// TIA Portal project "CMoLibrary_Dev" (V20)

(* hardware
DEVICE "S7-1500/ET200MP station_1"  S7-1500 station
   slot 0: "Rail_0"  Rack  6ES7 590-1***0-0AA0
   slot 1: "PLC_1"  CPU 1516-3 PN/DP  6ES7 516-3AN00-0AB0  V1.8
      slot 3: "CPU display_1"  6ES7591-1BA00-0AA0
      slot 32768: "PROFINET interface_1"  X1
         slot 32769: "Port_1"  X1 P1
         slot 32770: "Port_2"  X1 P2
      slot 33024: "PROFINET interface_2"  X2
         slot 33025: "Port_1"  X2 P1
      slot 33280: "DP interface_1"  X3
*)

// ===== PLC "PLC_1"  CPU 1516-3 PN/DP =====

TYPE "CMoDateTime"
   STRUCT
      RawDateTime : Array[0..6] of DInt;   // Platform-native wall clock data
      Year : DInt := 0;
      Month : DInt := 0;   // 1-12
      Day : DInt := 0;   // 1-31
      Hour : DInt := 0;   // 0-23
      Minute : DInt := 0;   // 0-59
      Second : DInt := 0;   // 0-59
      MicroSecond : DInt := 0;   // 0-999999
      IsLocal : Bool := false;   // TRUE = local time, FALSE = UTC
   END_STRUCT;
END_TYPE

TYPE "CMoDateTimeString"
   STRUCT
      TimeString : String[16];   // HH:MM:SS
      DateString : String[16];   // YYYY-MM-DD
      HMIString : String[32];   // YYYY-MM-DD HH:MM:SS
   END_STRUCT;
END_TYPE

TYPE "CMoHALDigitalInput"
   STRUCT
      Input : Bool := false;   // Raw hardware input (written by device driver)
      QualityInput : Bool := false;   // Hardware health from module status (TRUE = good)
      SimInput : Bool := false;   // Simulation input (written by twin/test)
      EnableSimulation : Bool := false;   // Enable simulation for this point
      SimulationIsActive : Bool := false;   // Computed: EnableSimulation AND Framework.SimulationEnabled
      HandValue : Bool := false;   // Manual override value (set from HMI)
      EnableHand : Bool := false;   // Enable hand mode for this point
      HandIsActive : Bool := false;   // Computed: EnableHand AND Framework.MaintenanceEnabled
      Value : Bool := false;   // THE OUTPUT: conditioned, filtered, mode-selected result
      Inverted : Bool := false;   // Invert input polarity
      BadQualityValue : Bool := false;   // Value to use when quality is bad (safe state)
      EnableDelay : Bool := false;   // Enable debounce filtering
      IsSpare : Bool := false;   // Mark as spare (bypasses quality, forces sim)
      InFilterOnTimeMsec : DInt := 0;   // On-delay debounce (milliseconds)
      InFilterOffTimeMsec : DInt := 0;   // Off-delay debounce (milliseconds)
      PointQuality : Bool := false;   // Computed quality (good if hw OK or sim active)
      RisingEdge : Bool := false;   // One-shot pulse on Value 0 to 1
      FallingEdge : Bool := false;   // One-shot pulse on Value 1 to 0
      "Name" : String[28];   // Human-readable tag name for HMI display
   END_STRUCT;
END_TYPE

TYPE "CMoHALDigitalOutput"
   STRUCT
      Output : Bool := false;   // Physical output (written by FB to hardware)
      QualityInput : Bool := false;   // Hardware health (TRUE = good)
      SimOutput : Bool := false;   // Shadow output for twin consumption during sim
      EnableSimulation : Bool := false;   // Enable simulation for this point
      SimulationIsActive : Bool := false;   // Computed: EnableSimulation AND Framework.SimulationEnabled
      HandValue : Bool := false;   // Manual override value (set from HMI)
      EnableHand : Bool := false;   // Enable hand mode for this point
      HandIsActive : Bool := false;   // Computed: EnableHand AND Framework.MaintenanceEnabled
      Value : Bool := false;   // Business logic command
      Inverted : Bool := false;   // Invert output polarity
      BadQualityValue : Bool := false;   // Value when quality is bad (safe state)
      IsSpare : Bool := false;   // Mark as spare
      PointQuality : Bool := false;   // Computed quality
      "Name" : String[28];   // Human-readable tag name
   END_STRUCT;
END_TYPE

TYPE "CMoInterlock"
   STRUCT
      PointCount : Int := 4;   // Number of active conditions (1-16)
      Condition : Array[0..15] of Bool;   // Condition inputs (set by business logic each scan)
      Bypass : Array[0..15] of Bool;   // Per-condition bypass (set from HMI)
      OK : Bool := false;   // All active conditions met (or bypassed)
      InBypass : Bool := false;   // At least one condition is bypassed
      BypassAlarm : Bool := false;   // Alarm: operating with bypassed conditions
      FirstOut : Int := -1;   // Index of first condition to drop (-1 = none)
      ConditionMet : Array[0..15] of Bool;   // Condition OR its bypass
      ConditionFaulted : Array[0..15] of Bool;   // Failed AND not bypassed
      "Name" : String[28];   // Interlock name
      ConditionName : Array[0..15] of String[28];   // Per-condition labels
   END_STRUCT;
END_TYPE

TYPE "CMoFramework"
   STRUCT
      AnyAudibleOn : Bool := false;   // At least one alarm has audible active
      AnyAudibleOnLastScan : Bool := false;   // Scratch accumulator
      AnyAlarmActive : Bool := false;   // At least one alarm active
      AnyAlarmActiveLastScan : Bool := false;   // Scratch accumulator
      AnyWarningActive : Bool := false;   // At least one warning-severity alarm
      AnyWarningActiveLastScan : Bool := false;   // Scratch accumulator
      AnyFaultActive : Bool := false;   // At least one fault-severity alarm
      AnyFaultActiveLastScan : Bool := false;   // Scratch accumulator
      AnyCriticalActive : Bool := false;   // At least one critical-severity alarm
      AnyCriticalActiveLastScan : Bool := false;   // Scratch accumulator
      AnySimulationOn : Bool := false;   // At least one I/O in simulation mode
      AnySimulationOnLastScan : Bool := false;   // Scratch accumulator
      AnyHandOn : Bool := false;   // At least one I/O in hand mode
      AnyHandOnLastScan : Bool := false;   // Scratch accumulator
      SilenceCmd : Bool := false;   // HMI silence button (momentary)
      GlobalAlmRstCmd : Bool := false;   // HMI global alarm reset (momentary)
      GlobalAlmRstEn : Bool := false;   // Enable global alarm reset
      SimulationEnabled : Bool := false;   // Master simulation enable
      EmulationEnabled : Bool := false;   // Running on emulated controller
      MaintenanceEnabled : Bool := false;   // Enables Hand mode
      Tick100ms : Bool := false;   // Pulse TRUE for one scan every 100ms
      Tick1s : Bool := false;   // Pulse TRUE for one scan every 1s
      Tick10s : Bool := false;   // Pulse TRUE for one scan every 10s
      Blink100ms : Bool := false;   // 100ms on/off blinker
      Blink250ms : Bool := false;   // 250ms on/off blinker
      Blink500ms : Bool := false;   // 500ms on/off blinker
      Blink1s : Bool := false;   // 1s on/off blinker
      Blink2s : Bool := false;   // 2s on/off blinker
      InhibitAlarms : Bool := false;   // Corporate alarm inhibit
      AlwaysTrue : Bool := false;   // Constant TRUE
      AlwaysFalse : Bool := false;   // Constant FALSE
      ApplicationCount : DInt := 0;   // Number of AOI instances registered
      AlarmCount : Int := 0;   // Current active alarm count
      TempAlarmCount : Int := 0;   // Scratch accumulator
      FreeRunningTimer : DInt := 0;   // Free-running ms counter
      LastRandomSeed : DInt := 0;   // Seed for random number generator
      Random : Real := 0.0;   // Current random number 0.0-1.0
      CycleTime : Real := 0.0;   // Last scan time (milliseconds)
      InhibitAlarmGroups : Array[0..15] of DWord;   // Per-group alarm inhibit (512 groups)
      CurrentUTCDateTime : "CMoDateTime";   // Current UTC time
      CurrentLocalDateTime : "CMoDateTime";   // Current local time
      CurrentUTCString : "CMoDateTimeString";   // UTC time formatted strings
      CurrentLocalString : "CMoDateTimeString";   // Local time formatted strings
      NotUsedDI : "CMoHALDigitalInput";   // Spare DI HAL instance
      NotUsedDO : "CMoHALDigitalOutput";   // Spare DO HAL instance
      ModuleStatusMinInterval : DInt := 5000;   // ms between module checks
      ModuleStatusRandomDistribution : DInt := 2000;   // ms random spread for check timing
      ModuleStatusGraceTime : DInt := 30000;   // ms before declaring module lost
   END_STRUCT;
END_TYPE

DATA_BLOCK "GVL"   // DB1
{ S7_Optimized_Access := 'TRUE' }
VERSION : 0.1
   VAR
      Framework : "CMoFramework";
      DI_PartPresent : "CMoHALDigitalInput";
      DI_GuardClosed : "CMoHALDigitalInput";
      DO_MotorRun : "CMoHALDigitalOutput";
      Interlock_Motor : "CMoInterlock";
      SimPartPresent : Bool;
      SimGuardClosed : Bool;
      saveStart : Bool;
      startDate : "CMoDateTime";
      saveEnd : Bool;
      endDate : "CMoDateTime";
   END_VAR
BEGIN
END_DATA_BLOCK

DATA_BLOCK "fbGuardClosed"   // DB2
{ S7_Optimized_Access := 'TRUE' }
VERSION : 0.1
// stored: InstanceOfName CMoDigitalInput
"CMoDigitalInput"
BEGIN
END_DATA_BLOCK

DATA_BLOCK "fbInterlock"   // DB3
{ S7_Optimized_Access := 'TRUE' }
VERSION : 0.1
// stored: InstanceOfName CMoEvalInterlock
"CMoEvalInterlock"
BEGIN
END_DATA_BLOCK

DATA_BLOCK "fbPartPresent"   // DB4
{ S7_Optimized_Access := 'TRUE' }
VERSION : 0.1
// stored: InstanceOfName CMoDigitalInput
"CMoDigitalInput"
BEGIN
END_DATA_BLOCK

DATA_BLOCK "fbMainRoutine"   // DB5
{ S7_Optimized_Access := 'TRUE' }
VERSION : 0.1
// stored: InstanceOfName CMoMainRuntime
"CMoMainRuntime"
BEGIN
END_DATA_BLOCK

DATA_BLOCK "fbMotorRun"   // DB6
{ S7_Optimized_Access := 'TRUE' }
VERSION : 0.1
// stored: InstanceOfName CMoDigitalOutput
"CMoDigitalOutput"
BEGIN
END_DATA_BLOCK

DATA_BLOCK "CMoDiffTime_DB"   // DB7
{ S7_Optimized_Access := 'TRUE' }
VERSION : 0.1
// stored: InstanceOfName CMoDiffTime
"CMoDiffTime"
BEGIN
END_DATA_BLOCK

FUNCTION_BLOCK "CMoRandom"   // FB1, SCL
{ S7_Optimized_Access := 'TRUE' }
VERSION : 0.1
   VAR_INPUT
      Seed : DInt := 48271;
   END_VAR
   VAR_OUTPUT
      Out : Real;
      NewSeed : DInt;
   END_VAR
BEGIN

   // =============================================================================
   // CMoRandom â€” Random Number Generator
   // CMo Library v1.0
   // =============================================================================
   // Park-Miller linear congruential generator.
   // Outputs a REAL between 0.0 and 1.0.
   //
   // Feed Seed from Framework.LastRandomSeed, write NewSeed back after call.
   // Called internally by CMoMainRuntime every scan.
   //
   // Usage:
   //   fbRandom(Seed := Framework.LastRandomSeed);
   //   Framework.Random := fbRandom.Out;
   //   Framework.LastRandomSeed := fbRandom.NewSeed;
   // =============================================================================

   // Ensure positive seed
   IF #Seed <= 0 THEN
       #Seed := 1;
   END_IF;

   // Park-Miller LCG: next = (seed * 16807) MOD 2147483647
   #NewSeed := (#Seed MOD 127773) * 16807 - (#Seed / 127773) * 2836;
   IF #NewSeed <= 0 THEN
       #NewSeed := #NewSeed + 2147483647;
   END_IF;

   #Out := DINT_TO_REAL(#NewSeed) / 2147483647.0;
END_FUNCTION_BLOCK

FUNCTION_BLOCK "CMoGetLocalDateTime"   // FB2, SCL
{ S7_Optimized_Access := 'TRUE' }
VERSION : 0.1
   VAR_IN_OUT
      DateTime : "CMoDateTime";
   END_VAR
   VAR_TEMP
      dtlNow : DTL;
      retVal : Int;
   END_VAR
BEGIN

   // =============================================================================
   // CMoGetLocalDateTime â€” Read Local System Time (Siemens)
   // CMo Library v1.0
   // =============================================================================
   // Reads the local system time using RD_LOC_T and parses DTL fields
   // into CMoDateTime.
   //
   // Must be called cyclically. Called internally by CMoMainRuntime.
   //
   // Usage:
   //   fbLocal(DateTime := Framework.CurrentLocalDateTime);
   // =============================================================================

   #retVal := RD_LOC_T(#dtlNow);

   IF #retVal <= 1 THEN
       #DateTime.Year := INT_TO_DINT(#dtlNow.YEAR);
       #DateTime.Month := USINT_TO_DINT(#dtlNow.MONTH);
       #DateTime.Day := USINT_TO_DINT(#dtlNow.DAY);
       #DateTime.Hour := USINT_TO_DINT(#dtlNow.HOUR);
       #DateTime.Minute := USINT_TO_DINT(#dtlNow.MINUTE);
       #DateTime.Second := USINT_TO_DINT(#dtlNow.SECOND);
       #DateTime.MicroSecond := UDINT_TO_DINT(#dtlNow.NANOSECOND / 1000);
       #DateTime.IsLocal := TRUE;
   END_IF;
END_FUNCTION_BLOCK

FUNCTION_BLOCK "CMoGetUTCDateTime"   // FB3, SCL
{ S7_Optimized_Access := 'TRUE' }
VERSION : 0.1
   VAR_IN_OUT
      DateTime : "CMoDateTime";
   END_VAR
   VAR_TEMP
      dtlNow : DTL;
      retVal : Int;
   END_VAR
BEGIN

   // =============================================================================
   // CMoGetUTCDateTime â€” Read UTC System Time (Siemens)
   // CMo Library v1.0
   // =============================================================================
   // Reads the UTC system time using RD_SYS_T and parses DTL fields
   // into CMoDateTime.
   //
   // RD_SYS_T returns UTC on S7-1500.
   // Must be called cyclically. Called internally by CMoMainRuntime.
   //
   // Usage:
   //   fbUTC(DateTime := Framework.CurrentUTCDateTime);
   // =============================================================================

   #retVal := RD_SYS_T(#dtlNow);

   IF #retVal = 0 THEN
       #DateTime.Year := INT_TO_DINT(#dtlNow.YEAR);
       #DateTime.Month := USINT_TO_DINT(#dtlNow.MONTH);
       #DateTime.Day := USINT_TO_DINT(#dtlNow.DAY);
       #DateTime.Hour := USINT_TO_DINT(#dtlNow.HOUR);
       #DateTime.Minute := USINT_TO_DINT(#dtlNow.MINUTE);
       #DateTime.Second := USINT_TO_DINT(#dtlNow.SECOND);
       #DateTime.MicroSecond := UDINT_TO_DINT(#dtlNow.NANOSECOND / 1000);
       #DateTime.IsLocal := FALSE;
   END_IF;
END_FUNCTION_BLOCK

FUNCTION_BLOCK "CMoElapsedTime"   // FB4, SCL
{ S7_Optimized_Access := 'TRUE' }
VERSION : 0.1
   VAR_INPUT
      Start : Bool;
      Stop : Bool;
      Reset : Bool;
   END_VAR
   VAR_OUTPUT
      ElapsedMs : Real;
      Running : Bool;
   END_VAR
   VAR
      PrevStart : Bool;
      PrevStop : Bool;
      tmRun : TON_TIME;
      Capturing : Bool;
   END_VAR
BEGIN

   // =============================================================================
   // CMoElapsedTime â€” Elapsed Time Measurement
   // CMo Library v1.0
   // =============================================================================
   // Measures elapsed time between Start and Stop rising edges.
   // Uses a TON timer internally for millisecond-resolution measurement.
   // Live readout available via ElapsedMs while Running is TRUE.
   //
   // Usage:
   //   myTimer(Start := TRUE);       // Begin measurement
   //   // ... code or scans pass ...
   //   myTimer(Stop := TRUE);        // End measurement
   //   result := myTimer.ElapsedMs;  // Read duration in ms
   //   myTimer(Reset := TRUE);       // Clear for next use
   // =============================================================================

   // Reset: clear everything
   IF #Reset THEN
       #ElapsedMs := 0.0;
       #Running := FALSE;
       #Capturing := FALSE;
       RETURN;
   END_IF;

   // Start on rising edge
   IF #Start AND NOT #PrevStart THEN
       #Capturing := TRUE;
       #Running := TRUE;
       #tmRun(IN := FALSE,
              PT := T#24D);
   END_IF;
   #PrevStart := #Start;

   // Accumulate while running
   IF #Capturing THEN
       #tmRun(IN := TRUE,
              PT := T#24D);
       #ElapsedMs := DINT_TO_REAL(TIME_TO_DINT(#tmRun.ET));
   END_IF;

   // Stop on rising edge
   IF #Stop AND NOT #PrevStop AND #Capturing THEN
       #ElapsedMs := DINT_TO_REAL(TIME_TO_DINT(#tmRun.ET));
       #Capturing := FALSE;
       #Running := FALSE;
   END_IF;
   #PrevStop := #Stop;
END_FUNCTION_BLOCK

FUNCTION_BLOCK "CMoDateTimeToString"   // FB5, SCL
{ S7_Optimized_Access := 'TRUE' }
VERSION : 0.1
   VAR_INPUT
      DateTime : "CMoDateTime";
   END_VAR
   VAR_IN_OUT
      DateTimeString : "CMoDateTimeString";
   END_VAR
   VAR_TEMP
      sYear : String[5];
      sMonth : String[3];
      sDay : String[3];
      sHour : String[3];
      sMinute : String[3];
      sSecond : String[3];
      sTemp : String[40];
   END_VAR
BEGIN
   // =============================================================================
   // CMoDateTimeToString — Format DateTime for HMI Display
   // CMo Library v1.0
   // =============================================================================
   // Converts CMoDateTime fields into zero-padded human-readable strings:
   //   TimeString: "HH:MM:SS"
   //   DateString: "YYYY-MM-DD"
   //   HMIString:  "YYYY-MM-DD HH:MM:SS"
   //
   // Siemens DINT_TO_STRING prepends a '+' sign. DELETE strips it.
   //
   // Usage:
   //   fbFmt(DateTime := myTime, DateTimeString := myStrings);
   // =============================================================================

   // Convert and strip leading '+'
   #sYear := DELETE(IN := DINT_TO_STRING(#DateTime.Year), L := 1, P := 1);

   IF #DateTime.Month < 10 THEN
       #sMonth := CONCAT(IN1 := '0', IN2 := DELETE(IN := DINT_TO_STRING(#DateTime.Month), L := 1, P := 1));
   ELSE
       #sMonth := DELETE(IN := DINT_TO_STRING(#DateTime.Month), L := 1, P := 1);
   END_IF;

   IF #DateTime.Day < 10 THEN
       #sDay := CONCAT(IN1 := '0', IN2 := DELETE(IN := DINT_TO_STRING(#DateTime.Day), L := 1, P := 1));
   ELSE
       #sDay := DELETE(IN := DINT_TO_STRING(#DateTime.Day), L := 1, P := 1);
   END_IF;

   IF #DateTime.Hour < 10 THEN
       #sHour := CONCAT(IN1 := '0', IN2 := DELETE(IN := DINT_TO_STRING(#DateTime.Hour), L := 1, P := 1));
   ELSE
       #sHour := DELETE(IN := DINT_TO_STRING(#DateTime.Hour), L := 1, P := 1);
   END_IF;

   IF #DateTime.Minute < 10 THEN
       #sMinute := CONCAT(IN1 := '0', IN2 := DELETE(IN := DINT_TO_STRING(#DateTime.Minute), L := 1, P := 1));
   ELSE
       #sMinute := DELETE(IN := DINT_TO_STRING(#DateTime.Minute), L := 1, P := 1);
   END_IF;

   IF #DateTime.Second < 10 THEN
       #sSecond := CONCAT(IN1 := '0', IN2 := DELETE(IN := DINT_TO_STRING(#DateTime.Second), L := 1, P := 1));
   ELSE
       #sSecond := DELETE(IN := DINT_TO_STRING(#DateTime.Second), L := 1, P := 1);
   END_IF;

   // Build TimeString: "HH:MM:SS"
   #sTemp := CONCAT(IN1 := #sHour, IN2 := ':');
   #sTemp := CONCAT(IN1 := #sTemp, IN2 := #sMinute);
   #sTemp := CONCAT(IN1 := #sTemp, IN2 := ':');
   #sTemp := CONCAT(IN1 := #sTemp, IN2 := #sSecond);
   #DateTimeString.TimeString := #sTemp;

   // Build DateString: "YYYY-MM-DD"
   #sTemp := CONCAT(IN1 := #sYear, IN2 := '-');
   #sTemp := CONCAT(IN1 := #sTemp, IN2 := #sMonth);
   #sTemp := CONCAT(IN1 := #sTemp, IN2 := '-');
   #sTemp := CONCAT(IN1 := #sTemp, IN2 := #sDay);
   #DateTimeString.DateString := #sTemp;

   // Build HMIString: "YYYY-MM-DD HH:MM:SS"
   #sTemp := CONCAT(IN1 := #DateTimeString.DateString, IN2 := ' ');
   #sTemp := CONCAT(IN1 := #sTemp, IN2 := #DateTimeString.TimeString);
   #DateTimeString.HMIString := #sTemp;
END_FUNCTION_BLOCK

FUNCTION_BLOCK "CMoDiffTime"   // FB6, SCL
{ S7_Optimized_Access := 'TRUE' }
VERSION : 0.1
   VAR_INPUT
      StartTime : "CMoDateTime";
      EndTime : "CMoDateTime";
   END_VAR
   VAR_OUTPUT
      Result : "CMoDateTime";
      TotalSeconds : DInt;
      TotalMicroseconds : DInt;
   END_VAR
   VAR_TEMP
      Borrow : DInt;
      Diff : DInt;
      "a" : DInt;
      y : DInt;
      "m" : DInt;
      jdnStart : DInt;
      jdnEnd : DInt;
      diffDays : DInt;
      diffUs : DInt;
      diffSec : DInt;
      diffMin : DInt;
      diffHr : DInt;
   END_VAR
BEGIN
   // =============================================================================
   // CMoDiffTime — DateTime Subtraction via Julian Day Number
   // CMo Library v1.0
   // =============================================================================
   // Computes (EndTime - StartTime) using Julian Day Number conversion.
   // Converts both dates to JDN (integer day count), subtracts, then
   // handles sub-day time remainder with borrow propagation.
   //
   // This is mathematically correct for all valid dates regardless of
   // month lengths, leap years, or century boundaries.
   //
   // Usage:
   //   fbDiff(StartTime := tStart, EndTime := tEnd);
   //   elapsed := fbDiff.TotalSeconds;
   // =============================================================================

   // JDN for StartTime
   #a := (14 - #StartTime.Month) / 12;
   #y := #StartTime.Year + 4800 - #a;
   #m := #StartTime.Month + 12 * #a - 3;
   #jdnStart := #StartTime.Day + (153 * #m + 2) / 5 + 365 * #y + #y / 4 - #y / 100 + #y / 400 - 32045;

   // JDN for EndTime
   #a := (14 - #EndTime.Month) / 12;
   #y := #EndTime.Year + 4800 - #a;
   #m := #EndTime.Month + 12 * #a - 3;
   #jdnEnd := #EndTime.Day + (153 * #m + 2) / 5 + 365 * #y + #y / 4 - #y / 100 + #y / 400 - 32045;

   // Day difference
   #diffDays := #jdnEnd - #jdnStart;

   // Sub-day difference with borrow propagation
   #diffUs := #EndTime.MicroSecond - #StartTime.MicroSecond;
   IF #diffUs < 0 THEN
       #diffUs := #diffUs + 1000000;
       #diffSec := -1;
   ELSE
       #diffSec := 0;
   END_IF;

   #diffSec := #diffSec + #EndTime.Second - #StartTime.Second;
   IF #diffSec < 0 THEN
       #diffSec := #diffSec + 60;
       #diffMin := -1;
   ELSE
       #diffMin := 0;
   END_IF;

   #diffMin := #diffMin + #EndTime.Minute - #StartTime.Minute;
   IF #diffMin < 0 THEN
       #diffMin := #diffMin + 60;
       #diffHr := -1;
   ELSE
       #diffHr := 0;
   END_IF;

   #diffHr := #diffHr + #EndTime.Hour - #StartTime.Hour;
   IF #diffHr < 0 THEN
       #diffHr := #diffHr + 24;
       #diffDays := #diffDays - 1;
   END_IF;

   // Populate result
   #Result.Year := 0;
   #Result.Month := 0;
   #Result.Day := #diffDays;
   #Result.Hour := #diffHr;
   #Result.Minute := #diffMin;
   #Result.Second := #diffSec;
   #Result.MicroSecond := #diffUs;
   #Result.IsLocal := FALSE;

   // Convenience totals
   #TotalSeconds := #diffSec + (#diffMin * 60) + (#diffHr * 3600) + (#diffDays * 86400);
   #TotalMicroseconds := #diffUs;
END_FUNCTION_BLOCK

FUNCTION_BLOCK "CMoAlarm"   // FB7, SCL
{ S7_Optimized_Access := 'TRUE' }
VERSION : 0.1
   VAR_INPUT
      Trigger : Bool;
      EnableAlarm : Bool := TRUE;
      AlarmOnTrue : Bool := TRUE;
      AutoReset : Bool;
      Delay : DInt;
      GroupNo : DInt;
      ID : Int;
      IsWarning : Bool;
      IsFault : Bool;
      IsCritical : Bool;
      EnableAudio : Bool;
      SystemResetEnable : Bool := TRUE;
      Inhibit : Bool;
      CountPreset : DInt;
   END_VAR
   VAR_OUTPUT
      AlarmActive : Bool;
      InhibitActive : Bool;
      AlarmCount : DInt;
      CountExceeded : Bool;
      AlarmSilenced : Bool;
   END_VAR
   VAR_IN_OUT
      Framework : "CMoFramework";
      CountReset : Bool;
      Reset : Bool;
   END_VAR
   VAR
      AlarmTimer : TON_TIME;
      IntGroupNo : DInt;
      IntID : DInt;
      IntReset : Bool;
      TriggerCondition : Bool;
      PrevAlarmActive : Bool;
      GroupWord : DInt;
      GroupBit : DInt;
   END_VAR
BEGIN

   // =============================================================================
   // CMoAlarm â€” Alarm Monitor
   // CMo Library v1.0
   // =============================================================================
   // Monitors a trigger condition and manages alarm lifecycle.
   // Supports configurable trigger polarity, delay before activation,
   // auto/manual reset, occurrence counting with threshold,
   // severity classification (Warning/Fault/Critical), group-based
   // inhibit, and HMI silencing.
   //
   // Usage:
   //   fbAlarm(
   //       Framework := GVL.Framework,
   //       Trigger := SomeCondition,
   //       ID := 100,
   //       Delay := 2000,
   //       IsFault := TRUE
   //   );
   // =============================================================================

   // Clamp group and ID
   IF #GroupNo >= 0 AND #GroupNo <= 511 THEN
       #IntGroupNo := #GroupNo;
   ELSE
       #IntGroupNo := 0;
   END_IF;

   IF #ID >= 1 AND #ID <= 9023 THEN
       #IntID := #ID;
   ELSE
       #IntID := 0;
   END_IF;

   #GroupWord := #IntGroupNo / 32;
   #GroupBit := #IntGroupNo MOD 32;

   // Count reset
   IF #CountReset THEN
       #AlarmCount := 0;
       #CountReset := FALSE;
   END_IF;

   // Inhibit evaluation
   #InhibitActive := NOT #EnableAlarm
   OR #Inhibit
   OR #Framework.InhibitAlarms;
   IF NOT #InhibitActive AND (#Framework.InhibitAlarmGroups[#GroupWord] AND SHL(IN := DWORD#1, N := DINT_TO_INT(#GroupBit))) <> 0 THEN
       #InhibitActive := TRUE;
   END_IF;

   // Composite reset
   #IntReset := #AutoReset
   OR #Reset
   OR (#SystemResetEnable AND #Framework.GlobalAlmRstEn AND #Framework.GlobalAlmRstCmd);

   // Trigger polarity
   IF #AlarmOnTrue THEN
       #TriggerCondition := #Trigger;
   ELSE
       #TriggerCondition := NOT #Trigger;
   END_IF;

   // Alarm activation with delay
   IF #IntID <> 0 THEN
       #AlarmTimer(
                   IN := (NOT #InhibitActive AND #TriggerCondition) OR (#AlarmActive AND NOT #IntReset),
                   PT := DINT_TO_TIME(#Delay)
       );
       #AlarmActive := #AlarmTimer.Q;
   ELSE
       #AlarmActive := FALSE;
   END_IF;

   // Count activations (rising edge)
   IF #AlarmActive AND NOT #PrevAlarmActive THEN
       #AlarmCount := #AlarmCount + 1;
   END_IF;

   // Silence
   IF #AlarmActive THEN
       IF #Framework.SilenceCmd OR #AlarmSilenced THEN
           #AlarmSilenced := TRUE;
       END_IF;
   ELSE
       #AlarmSilenced := FALSE;
   END_IF;

   // Roll up into Framework
   IF #AlarmActive THEN
       #Framework.TempAlarmCount := #Framework.TempAlarmCount + 1;
       #Framework.AnyAlarmActiveLastScan := TRUE;

       IF NOT #AlarmSilenced THEN
           IF #EnableAudio THEN
               #Framework.AnyAudibleOnLastScan := TRUE;
           END_IF;
           IF #IsWarning THEN
               #Framework.AnyWarningActiveLastScan := TRUE;
           END_IF;
           IF #IsFault THEN
               #Framework.AnyFaultActiveLastScan := TRUE;
           END_IF;
           IF #IsCritical THEN
               #Framework.AnyCriticalActiveLastScan := TRUE;
           END_IF;
       END_IF;
   END_IF;

   // Count threshold
   #CountExceeded := (#CountPreset > 0) AND (#AlarmCount >= #CountPreset);

   // Clear manual reset
   #Reset := FALSE;

   // Previous state
   #PrevAlarmActive := #AlarmActive;
END_FUNCTION_BLOCK

FUNCTION_BLOCK "CMoDigitalInput"   // FB8, SCL
{ S7_Optimized_Access := 'TRUE' }
VERSION : 0.1
   VAR_INPUT
      DeviceInput : Bool;
      QualityInput : Bool;
   END_VAR
   VAR_IN_OUT
      HAL : "CMoHALDigitalInput";
      Framework : "CMoFramework";
   END_VAR
   VAR
      ConditionedInput : Bool;
      DebouncedValue : Bool;
      OnDelayTimer : TON_TIME;
      OffDelayTimer : TOF_TIME;
      PrevValue : Bool;
      FirstScan : Bool := TRUE;
      ReSync : Bool;
      NoFilterNeeded : Bool;
   END_VAR
BEGIN

   // =============================================================================
   // CMoDigitalInput â€” Digital Input Signal Conditioning
   // CMo Library v1.0
   // =============================================================================
   // Takes a raw hardware input and produces a conditioned .Value through:
   //   1. Mode determination (Normal / Simulation / Hand)
   //   2. Quality evaluation (hardware health, sim, spare)
   //   3. Mode selection + polarity inversion
   //   4. Debounce filtering (configurable on/off delay with resync)
   //   5. Hand value bumpless transfer
   //   6. Quality gating (bad quality -> configurable fallback)
   //   7. Edge detection (RisingEdge / FallingEdge one-shot pulses)
   //
   // Business logic reads .Value only. Never touch .Input, .SimInput,
   // .HandValue, or any plumbing directly.
   //
   // Usage:
   //   fbInput(
   //       HAL := GVL.MyInput,
   //       DeviceInput := Module1:I.Data[0],
   //       QualityInput := Module1_Status.Running,
   //       Framework := GVL.Framework
   //   );
   // =============================================================================

   // Mode determination
   #HAL.HandIsActive := #HAL.EnableHand AND #Framework.MaintenanceEnabled;
   IF #HAL.HandIsActive THEN
       #Framework.AnyHandOnLastScan := TRUE;
   END_IF;

   #HAL.SimulationIsActive := #HAL.EnableSimulation AND #Framework.SimulationEnabled;
   IF #HAL.SimulationIsActive THEN
       #Framework.AnySimulationOnLastScan := TRUE;
   END_IF;

   // Point quality
   IF #HAL.IsSpare THEN
       #HAL.PointQuality := TRUE;
   ELSIF #HAL.SimulationIsActive THEN
       #HAL.PointQuality := TRUE;
   ELSE
       #HAL.QualityInput := #QualityInput;
       #HAL.PointQuality := #QualityInput;
   END_IF;

   // Latch raw input
   #HAL.Input := #DeviceInput;

   // Mode selection + inversion
   IF #HAL.SimulationIsActive THEN
       IF #HAL.Inverted THEN
           #ConditionedInput := NOT #HAL.SimInput;
       ELSE
           #ConditionedInput := #HAL.SimInput;
       END_IF;
   ELSE
       IF #HAL.Inverted THEN
           #ConditionedInput := NOT #HAL.Input;
       ELSE
           #ConditionedInput := #HAL.Input;
       END_IF;
   END_IF;

   // Debounce filter
   IF NOT #HAL.EnableDelay THEN
       #DebouncedValue := #ConditionedInput;
       #ReSync := TRUE;
   ELSE
       IF #HAL.InFilterOnTimeMsec < 0 THEN
           #HAL.InFilterOnTimeMsec := 0;
       END_IF;
       IF #HAL.InFilterOffTimeMsec < 0 THEN
           #HAL.InFilterOffTimeMsec := 0;
       END_IF;

       #OnDelayTimer(
                     IN := #ConditionedInput OR (#OffDelayTimer.Q AND #OnDelayTimer.Q),
                     PT := DINT_TO_TIME(#HAL.InFilterOnTimeMsec)
       );

       #OffDelayTimer(
                      IN := #ConditionedInput,
                      PT := DINT_TO_TIME(#HAL.InFilterOffTimeMsec)
       );

       #NoFilterNeeded := (#ConditionedInput AND #OnDelayTimer.Q)
       OR (NOT #ConditionedInput AND NOT #OffDelayTimer.Q);

       IF #ReSync THEN
           IF (#DebouncedValue AND #OnDelayTimer.Q) OR
               (NOT #DebouncedValue AND NOT #OnDelayTimer.Q) THEN
               #ReSync := FALSE;
           END_IF;
       END_IF;

       IF #ReSync OR #HAL.IsSpare THEN
           #DebouncedValue := #ConditionedInput;
       ELSIF #OnDelayTimer.Q THEN
           #DebouncedValue := TRUE;
       ELSIF NOT #OffDelayTimer.Q THEN
           #DebouncedValue := FALSE;
       END_IF;
   END_IF;

   // Hand value tracking (bumpless transfer)
   IF NOT #HAL.HandIsActive THEN
       #HAL.HandValue := #HAL.Value;
   END_IF;

   // Final value with quality gating
   IF #HAL.PointQuality THEN
       IF #HAL.HandIsActive THEN
           #HAL.Value := #HAL.HandValue;
       ELSE
           #HAL.Value := #DebouncedValue;
       END_IF;
   ELSE
       #HAL.Value := #HAL.BadQualityValue;
   END_IF;

   // Edge detection
   IF #FirstScan THEN
       #PrevValue := #HAL.Value;
       #HAL.RisingEdge := FALSE;
       #HAL.FallingEdge := FALSE;
       #FirstScan := FALSE;
   ELSE
       #HAL.RisingEdge := #HAL.Value AND NOT #PrevValue;
       #HAL.FallingEdge := NOT #HAL.Value AND #PrevValue;
       #PrevValue := #HAL.Value;
   END_IF;
END_FUNCTION_BLOCK

FUNCTION_BLOCK "CMoDigitalOutput"   // FB9, SCL
{ S7_Optimized_Access := 'TRUE' }
VERSION : 0.1
   VAR_INPUT
      QualityInput : Bool;
   END_VAR
   VAR_OUTPUT
      DeviceOutput : Bool;
   END_VAR
   VAR_IN_OUT
      HAL : "CMoHALDigitalOutput";
      Framework : "CMoFramework";
   END_VAR
   VAR
      ConditionedOutput : Bool;
      OutputWithHand : Bool;
   END_VAR
BEGIN

   // =============================================================================
   // CMoDigitalOutput â€” Digital Output Signal Conditioning
   // CMo Library v1.0
   // =============================================================================
   // Takes .Value written by business logic and produces a conditioned
   // physical output through:
   //   1. Mode determination (Normal / Simulation / Hand)
   //   2. Quality evaluation (hardware health, sim, spare)
   //   3. Polarity inversion
   //   4. Hand value bumpless transfer
   //   5. Hand mode selection
   //   6. Simulation gating (suppress physical output, capture to .SimOutput)
   //
   // In simulation mode: DeviceOutput is suppressed. The digital twin
   // reads .SimOutput to see what business logic commanded.
   //
   // Usage:
   //   fbOutput(
   //       HAL := GVL.MyOutput,
   //       QualityInput := Module2_Status.Running,
   //       Framework := GVL.Framework
   //   );
   //   Module2:O.Data[0] := fbOutput.DeviceOutput;
   // =============================================================================

   // Mode determination
   #HAL.HandIsActive := #HAL.EnableHand AND #Framework.MaintenanceEnabled AND NOT #HAL.IsSpare;
   IF #HAL.HandIsActive THEN
       #Framework.AnyHandOnLastScan := TRUE;
   END_IF;

   #HAL.SimulationIsActive := #HAL.EnableSimulation AND #Framework.SimulationEnabled;
   IF #HAL.SimulationIsActive THEN
       #Framework.AnySimulationOnLastScan := TRUE;
   END_IF;

   // Point quality
   IF #HAL.IsSpare THEN
       #HAL.PointQuality := TRUE;
   ELSIF #HAL.SimulationIsActive THEN
       #HAL.PointQuality := TRUE;
   ELSE
       #HAL.QualityInput := #QualityInput;
       #HAL.PointQuality := #QualityInput;
   END_IF;

   // Inversion
   IF NOT #HAL.IsSpare THEN
       IF #HAL.Inverted THEN
           #ConditionedOutput := NOT #HAL.Value;
       ELSE
           #ConditionedOutput := #HAL.Value;
       END_IF;
   ELSE
       #ConditionedOutput := FALSE;
   END_IF;

   // Hand value tracking (bumpless transfer)
   IF NOT #HAL.HandIsActive THEN
       #HAL.HandValue := #HAL.Value;
   END_IF;

   // Hand mode selection
   IF #HAL.HandIsActive THEN
       #OutputWithHand := #HAL.HandValue;
   ELSE
       #OutputWithHand := #ConditionedOutput;
   END_IF;

   // Simulation gating
   IF #HAL.SimulationIsActive THEN
       #DeviceOutput := FALSE;
   ELSE
       #DeviceOutput := #OutputWithHand;
   END_IF;

   #HAL.SimOutput := #OutputWithHand;
   #HAL.Output := #DeviceOutput;
END_FUNCTION_BLOCK

FUNCTION_BLOCK "CMoEvalInterlock"   // FB10, SCL
{ S7_Optimized_Access := 'TRUE' }
VERSION : 0.1
   VAR_IN_OUT
      Ilk : "CMoInterlock";
   END_VAR
   VAR
      PrevOK : Bool;
   END_VAR
   VAR_TEMP
      i : Int;
      AllMet : Bool;
      AnyBypassed : Bool;
      FirstDropped : Int;
   END_VAR
BEGIN

   // =============================================================================
   // CMoEvalInterlock â€” Interlock Evaluation
   // CMo Library v1.0
   // =============================================================================
   // Evaluates up to 16 AND conditions with first-out tracking
   // and per-condition bypass. All active conditions must be TRUE
   // (or bypassed) for .OK to be TRUE.
   //
   // FirstOut latches the index of the first faulted condition on
   // the OK->NOT OK transition (root cause analysis from HMI).
   //
   // Usage:
   //   Ilk.Condition[0] := EStop.Value;
   //   Ilk.Condition[1] := GuardDoor.Value;
   //   fbInterlock(Ilk := MyInterlock);
   //   IF MyInterlock.OK THEN ... END_IF;
   // =============================================================================

   // Clamp PointCount
   IF #Ilk.PointCount < 1 THEN
       #Ilk.PointCount := 1;
   ELSIF #Ilk.PointCount > 16 THEN
       #Ilk.PointCount := 16;
   END_IF;

   // Evaluate each condition
   #AllMet := TRUE;
   #AnyBypassed := FALSE;
   #FirstDropped := -1;

   FOR #i := 0 TO #Ilk.PointCount - 1 DO
       #Ilk.ConditionMet[#i] := #Ilk.Condition[#i] OR #Ilk.Bypass[#i];
       #Ilk.ConditionFaulted[#i] := NOT #Ilk.Condition[#i] AND NOT #Ilk.Bypass[#i];

       IF #Ilk.Bypass[#i] THEN
           #AnyBypassed := TRUE;
       END_IF;

       IF #Ilk.ConditionFaulted[#i] AND #FirstDropped = -1 THEN
           #FirstDropped := #i;
       END_IF;

       IF NOT #Ilk.ConditionMet[#i] THEN
           #AllMet := FALSE;
       END_IF;
   END_FOR;

   // Clear unused conditions
   FOR #i := #Ilk.PointCount TO 15 DO
       #Ilk.ConditionMet[#i] := TRUE;
       #Ilk.ConditionFaulted[#i] := FALSE;
   END_FOR;

   // Outputs
   #PrevOK := #Ilk.OK;
   #Ilk.OK := #AllMet;
   #Ilk.InBypass := #AnyBypassed;
   #Ilk.BypassAlarm := #AnyBypassed;

   // FirstOut: latch on OK->NOT OK transition
   IF NOT #Ilk.OK AND #PrevOK THEN
       #Ilk.FirstOut := #FirstDropped;
   ELSIF #Ilk.OK THEN
       #Ilk.FirstOut := -1;
   END_IF;
END_FUNCTION_BLOCK

FUNCTION_BLOCK "CMoMainRuntime"   // FB11, SCL
{ S7_Optimized_Access := 'TRUE' }
VERSION : 0.1
   VAR_IN_OUT
      Framework : "CMoFramework";
   END_VAR
   VAR
      tmTick100ms : TON_TIME;
      tmTick1s : TON_TIME;
      tmTick10s : TON_TIME;
      tmBlink100ms : TON_TIME;
      tmBlink250ms : TON_TIME;
      tmBlink500ms : TON_TIME;
      tmBlink1s : TON_TIME;
      tmBlink2s : TON_TIME;
      bState100ms : Bool;
      bState250ms : Bool;
      bState500ms : Bool;
      bState1s : Bool;
      bState2s : Bool;
      fbGetLocal : "CMoGetLocalDateTime";
      fbGetUTC : "CMoGetUTCDateTime";
      fbLocalToStr : "CMoDateTimeToString";
      fbUTCToStr : "CMoDateTimeToString";
      fbScanTime : "CMoElapsedTime";
      bScanRunning : Bool;
      fbRandom : "CMoRandom";
   END_VAR
BEGIN

   // =============================================================================
   // CMoMainRuntime â€” System Heartbeat
   // CMo Library v1.0
   // =============================================================================
   // Call ONCE per scan, FIRST in the task. Responsible for:
   //   - Measuring scan cycle time (via CMoElapsedTime)
   //   - Generating tick timers (100ms, 1s, 10s)
   //   - Generating blinker signals (100ms, 250ms, 500ms, 1s, 2s)
   //   - Latching LastScan accumulators into final alarm/sim/hand rollups
   //   - Resetting LastScan accumulators for the new scan
   //   - Generating random number (via CMoRandom)
   //   - Updating local and UTC date/time with formatted strings
   //   - Setting constants (AlwaysTrue, AlwaysFalse)
   //   - Incrementing free-running timer
   //
   // The LastScan pattern:
   //   MainRuntime resets all *LastScan fields at start of scan.
   //   Individual CMoAlarm/CMoDigitalInput FBs SET them during the scan.
   //   MainRuntime copies LastScan -> final at the NEXT call.
   //   This eliminates execution order dependencies.
   //
   // Usage:
   //   fbRuntime(Framework := GVL.Framework);  // first line of MAIN
   // =============================================================================

   // Scan time measurement: stop previous, read result, start new
   IF #bScanRunning THEN
       #fbScanTime(Start := FALSE,
                   Stop := TRUE,
                   Reset := FALSE);
       #Framework.CycleTime := #fbScanTime.ElapsedMs;
       #fbScanTime(Start := FALSE,
                   Stop := FALSE,
                   Reset := TRUE);
       #fbScanTime(Start := TRUE,
                   Stop := FALSE,
                   Reset := FALSE);
   ELSE
       #fbScanTime(Start := TRUE,
                   Stop := FALSE,
                   Reset := FALSE);
       #bScanRunning := TRUE;
   END_IF;

   // Latch previous scan accumulators into final outputs
   #Framework.AnyAudibleOn := #Framework.AnyAudibleOnLastScan;
   #Framework.AnyAlarmActive := #Framework.AnyAlarmActiveLastScan;
   #Framework.AnyWarningActive := #Framework.AnyWarningActiveLastScan;
   #Framework.AnyFaultActive := #Framework.AnyFaultActiveLastScan;
   #Framework.AnyCriticalActive := #Framework.AnyCriticalActiveLastScan;
   #Framework.AnySimulationOn := #Framework.AnySimulationOnLastScan;
   #Framework.AnyHandOn := #Framework.AnyHandOnLastScan;
   #Framework.AlarmCount := #Framework.TempAlarmCount;

   // Reset scratch for this scan
   #Framework.AnyAudibleOnLastScan := FALSE;
   #Framework.AnyAlarmActiveLastScan := FALSE;
   #Framework.AnyWarningActiveLastScan := FALSE;
   #Framework.AnyFaultActiveLastScan := FALSE;
   #Framework.AnyCriticalActiveLastScan := FALSE;
   #Framework.AnySimulationOnLastScan := FALSE;
   #Framework.AnyHandOnLastScan := FALSE;
   #Framework.TempAlarmCount := 0;

   // Constants
   #Framework.AlwaysTrue := TRUE;
   #Framework.AlwaysFalse := FALSE;

   // Random number generator
   #fbRandom(Seed := #Framework.LastRandomSeed);
   #Framework.Random := #fbRandom.Out;
   #Framework.LastRandomSeed := #fbRandom.NewSeed;

   // Ticks: pulse TRUE for one scan at each interval
   #tmTick100ms(IN := TRUE,
                PT := T#100MS);
   #Framework.Tick100ms := #tmTick100ms.Q;
   IF #tmTick100ms.Q THEN
       #tmTick100ms(IN := FALSE,
                    PT := T#100MS);
   END_IF;

   #tmTick1s(IN := TRUE,
             PT := T#1S);
   #Framework.Tick1s := #tmTick1s.Q;
   IF #tmTick1s.Q THEN
       #tmTick1s(IN := FALSE,
                 PT := T#1S);
   END_IF;

   #tmTick10s(IN := TRUE,
              PT := T#10S);
   #Framework.Tick10s := #tmTick10s.Q;
   IF #tmTick10s.Q THEN
       #tmTick10s(IN := FALSE,
                  PT := T#10S);
   END_IF;

   // Blinkers: toggle state at each interval
   #tmBlink100ms(IN := TRUE,
                 PT := T#100MS);
   IF #tmBlink100ms.Q THEN
       #bState100ms := NOT #bState100ms;
       #tmBlink100ms(IN := FALSE,
                     PT := T#100MS);
   END_IF;
   #Framework.Blink100ms := #bState100ms;

   #tmBlink250ms(IN := TRUE,
                 PT := T#250MS);
   IF #tmBlink250ms.Q THEN
       #bState250ms := NOT #bState250ms;
       #tmBlink250ms(IN := FALSE,
                     PT := T#250MS);
   END_IF;
   #Framework.Blink250ms := #bState250ms;

   #tmBlink500ms(IN := TRUE,
                 PT := T#500MS);
   IF #tmBlink500ms.Q THEN
       #bState500ms := NOT #bState500ms;
       #tmBlink500ms(IN := FALSE,
                     PT := T#500MS);
   END_IF;
   #Framework.Blink500ms := #bState500ms;

   #tmBlink1s(IN := TRUE,
              PT := T#1S);
   IF #tmBlink1s.Q THEN
       #bState1s := NOT #bState1s;
       #tmBlink1s(IN := FALSE,
                  PT := T#1S);
   END_IF;
   #Framework.Blink1s := #bState1s;

   #tmBlink2s(IN := TRUE,
              PT := T#2S);
   IF #tmBlink2s.Q THEN
       #bState2s := NOT #bState2s;
       #tmBlink2s(IN := FALSE,
                  PT := T#2S);
   END_IF;
   #Framework.Blink2s := #bState2s;

   // Free-running timer
   #Framework.FreeRunningTimer := #Framework.FreeRunningTimer + 1;

   // Date/Time: read local and UTC, format strings
   #fbGetLocal(DateTime := #Framework.CurrentLocalDateTime);
   #fbGetUTC(DateTime := #Framework.CurrentUTCDateTime);

   #fbLocalToStr(
                 DateTime := #Framework.CurrentLocalDateTime,
                 DateTimeString := #Framework.CurrentLocalString
   );
   #fbUTCToStr(
               DateTime := #Framework.CurrentUTCDateTime,
               DateTimeString := #Framework.CurrentUTCString
   );
END_FUNCTION_BLOCK

ORGANIZATION_BLOCK "Main"   // OB1, FBD, ProgramCycle
TITLE = "Main Program Sweep (Cycle)"
{ S7_Optimized_Access := 'TRUE' }
VERSION : 0.1
   VAR_INPUT
      Initial_Call : Bool;   // Initial call of this OB
      Remanence : Bool;   // =True, if remanent data are available
   END_VAR
BEGIN

REGION Network 1
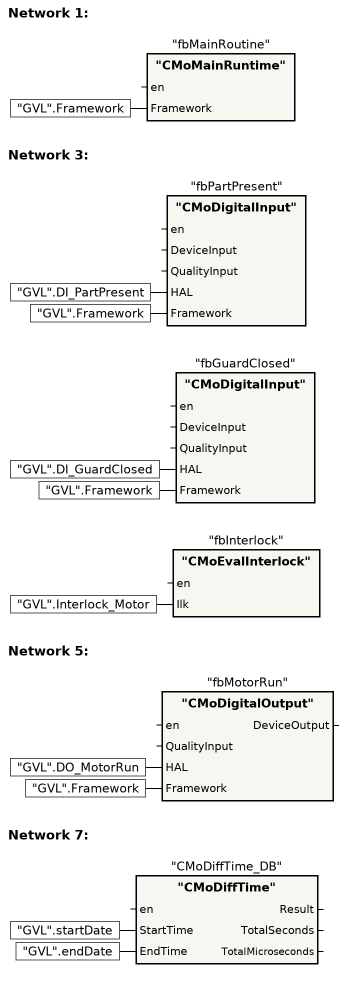
   "fbMainRoutine"(Framework := "GVL".Framework);   // "CMoMainRuntime"
END_REGION

REGION Network 2 (SCL)
   // Enable simulation globally
   "GVL".Framework.SimulationEnabled := TRUE;

   // --- Part Present sensor ---
   "GVL".DI_PartPresent.EnableSimulation := TRUE;
   "GVL".DI_PartPresent.SimInput := "GVL".SimPartPresent;
   "GVL".DI_PartPresent.Name := 'Part Present';

   // --- Guard Door sensor ---
   "GVL".DI_GuardClosed.EnableSimulation := TRUE;
   "GVL".DI_GuardClosed.SimInput := "GVL".SimGuardClosed;
   "GVL".DI_GuardClosed.Name := 'Guard Closed';

   // --- Interlock ---
   "GVL".Interlock_Motor.PointCount := 2;
   "GVL".Interlock_Motor.ConditionName[0] := 'Part Present';
   "GVL".Interlock_Motor.ConditionName[1] := 'Guard Closed';
   "GVL".Interlock_Motor.Condition[0] := "GVL".DI_PartPresent.Value;
   "GVL".Interlock_Motor.Condition[1] := "GVL".DI_GuardClosed.Value;
END_REGION

REGION Network 3
   "fbPartPresent"(HAL := "GVL".DI_PartPresent, Framework := "GVL".Framework);   // "CMoDigitalInput"
   "fbGuardClosed"(HAL := "GVL".DI_GuardClosed, Framework := "GVL".Framework);   // "CMoDigitalInput"
   "fbInterlock"(Ilk := "GVL".Interlock_Motor);   // "CMoEvalInterlock"
END_REGION

REGION Network 4 (SCL)
   // --- Business logic: .Value only ---
   "GVL".DO_MotorRun.EnableSimulation := TRUE;
   "GVL".DO_MotorRun.Value := "GVL".Interlock_Motor.OK;
   "GVL".DO_MotorRun.Name := 'Motor Run';
END_REGION

REGION Network 5
   "fbMotorRun"(HAL := "GVL".DO_MotorRun, Framework := "GVL".Framework);   // "CMoDigitalOutput"
END_REGION

REGION Network 6 (SCL)
   IF "GVL".saveStart = 1 THEN
       "GVL".startDate := "GVL".Framework.CurrentUTCDateTime;
   END_IF;
   IF "GVL".saveEnd = 1 THEN
       "GVL".endDate := "GVL".Framework.CurrentUTCDateTime;
   END_IF;
END_REGION

REGION Network 7
   "CMoDiffTime_DB"(StartTime := "GVL".startDate, EndTime := "GVL".endDate);   // "CMoDiffTime"
END_REGION
END_ORGANIZATION_BLOCK